(* IEC 61131-3 sources: codesys-framework/txt/application/WeVe IO (library)/DigitalOutput/FB_DigitalOutput, 2 files *)

(* ---- Output.prop.st ---- *)
PROPERTY Output : BOOL

// --- BEGIN IMPLEMENTATION ---

// ----------- SET -----------
VAR
END_VAR

// -- BEGIN IMPLEMENTATION SET --
_xOutputValue := Output;

// ----------- GET -----------
VAR
END_VAR

// -- BEGIN IMPLEMENTATION GET --
Output := _xOutputValue;

(* ---- SysPar.prop.st ---- *)
PROPERTY SysPar : SC_SystemParametersDigitalOutput

// --- BEGIN IMPLEMENTATION ---

// ----------- SET -----------
VAR
END_VAR

// -- BEGIN IMPLEMENTATION SET --
_scSysPar := SysPar;
